FUNCTION_BLOCK FB_SignalWatchdog
VAR_INPUT
	(* Input variables / Eingang Variablen *)
	bEnable					:BOOL;						(* Enable FB signal *)
	bIn						:BOOL;						(* Input signal *)
	tWatchdog				:TIME := t#0s;					(* Watchdog time *)
END_VAR
VAR_OUTPUT
	(* Output variables / Ausgang Variablen *)
	bOut					:BOOL;						(* Output signal *)
	bAlarm					:BOOL;						(* Alarm signal *)
END_VAR
VAR
	(* Enummerations *)

	(* Variables *)


	(* References *)

	(* Interfaces *)

	(* Instances *)
	tofWatchdog				:TOF;

END_VAR

IF NOT bEnable
THEN
	bOut := FALSE;
	bAlarm := FALSE;                       (* Alarm active *)
	
	tofWatchdog(
		IN := tofWatchdog.ET > t#0ms,
	         PT := t#0ms
	);
	
	tofWatchdog(IN := FALSE,
	             PT := t#0ms);

	RETURN;
END_IF;

tofWatchdog(					 (* Dealy input signal *)
	IN := bIn,
	PT := tWatchdog
);

bOut := tofWatchdog.Q;

bAlarm := NOT tofWatchdog.Q;                       (* Set alarm *)

END_FUNCTION_BLOCK

(* stored: Version 1.1.0.1, ProductVersion 3.1.4024.15
   POU FB_SignalWatchdog: Id {4fdbc35a-777b-4d30-88d6-1240b71a05ad}, SpecialFunc None *)
